screen "D_Rectangle_1" 1280x800
   TextField "Label_Static" at 6,86 size 148x16; Text 'Static'
   Rectangle "A_Range" at 158,4 size 100x50
      Appearance <- "D_Range"
   TextField "Label_A_Range" at 158,86 size 148x16; Text 'A_Range'
   Rectangle "A_Flash" at 310,4 size 100x50
      Appearance <- "D_Range"
   TextField "Label_A_Flash" at 310,86 size 148x16; Text 'A_Flash'
   Rectangle "A_Bit" at 462,4 size 100x50
      Appearance <- "D_Bool"
   TextField "Label_A_Bit" at 462,86 size 148x16; Text 'A_Bit'
   Rectangle "A_Bits" at 614,4 size 100x50
      Appearance <- "D_Bits"
   TextField "Label_A_Bits" at 614,86 size 148x16; Text 'A_Bits'
   Rectangle "V_Range" at 766,4 size 100x50
      Visibility <- "D_Range"
   TextField "Label_V_Range" at 766,86 size 148x16; Text 'V_Range'
   Rectangle "V_Bit" at 918,4 size 100x50
      Visibility <- "D_Vis"
   TextField "Label_V_Bit" at 918,86 size 148x16; Text 'V_Bit'
   Rectangle "M_H" at 1070,4 size 100x50
      HorizontalMovement <- "D_Pct"
   TextField "Label_M_H" at 1070,86 size 148x16; Text 'M_H'
   Rectangle "M_V" at 6,106 size 100x50
      VerticalMovement <- "D_Pct"
   TextField "Label_M_V" at 6,188 size 148x16; Text 'M_V'
   Rectangle "M_D" at 158,106 size 100x50
      DiagonalMovement <- "D_Pct"
   TextField "Label_M_D" at 158,188 size 148x16; Text 'M_D'
   Rectangle "M_Direct" at 310,106 size 100x50
      DirectMovement <- "D_X"
      DirectMovement <- "D_Y"
   TextField "Label_M_Direct" at 310,188 size 148x16; Text 'M_Direct'
   Rectangle "E_Range" at 462,106 size 100x50
      ObjectEnable <- "D_Range"
   TextField "Label_E_Range" at 462,188 size 148x16; Text 'E_Range'
   Rectangle "E_Bit" at 614,106 size 100x50
      ObjectEnable <- "D_En"
   TextField "Label_E_Bit" at 614,188 size 148x16; Text 'E_Bit'
   IOField "State" at 4,774 size 60x22; FormatPattern 9
      ProcessValue <- "D_State"
   Button "S1" at 70,774 size 40x22; TextOff 'S1'
      on Click: "SetS1"()
   Button "S2" at 114,774 size 40x22; TextOff 'S2'
      on Click: "SetS2"()
   Button "S3" at 158,774 size 40x22; TextOff 'S3'
      on Click: "SetS3"()
   Button "S4" at 202,774 size 40x22; TextOff 'S4'
      on Click: "SetS4"()
   Button "Next" at 1236,774 size 40x22; TextOff 'Next'
      on Click: ActivateScreen("D_TextField_1", 0)

screen "D_Slider_1" 1280x800
   Slider "Static" at 6,4 size 60x160; Caption 'SIMATIC'
   TextField "Label_Static" at 6,196 size 108x16; Text 'Static'
   Slider "A_Range" at 118,4 size 60x160; Caption 'SIMATIC'
      Appearance <- "D_Range"
   TextField "Label_A_Range" at 118,196 size 108x16; Text 'A_Range'
   Slider "A_Flash" at 230,4 size 60x160; Caption 'SIMATIC'
      Appearance <- "D_Range"
   TextField "Label_A_Flash" at 230,196 size 108x16; Text 'A_Flash'
   Slider "A_Bit" at 342,4 size 60x160; Caption 'SIMATIC'
      Appearance <- "D_Bool"
   TextField "Label_A_Bit" at 342,196 size 108x16; Text 'A_Bit'
   Slider "A_Bits" at 454,4 size 60x160; Caption 'SIMATIC'
      Appearance <- "D_Bits"
   TextField "Label_A_Bits" at 454,196 size 108x16; Text 'A_Bits'
   Slider "V_Range" at 566,4 size 60x160; Caption 'SIMATIC'
      Visibility <- "D_Range"
   TextField "Label_V_Range" at 566,196 size 108x16; Text 'V_Range'
   Slider "V_Bit" at 678,4 size 60x160; Caption 'SIMATIC'
      Visibility <- "D_Vis"
   TextField "Label_V_Bit" at 678,196 size 108x16; Text 'V_Bit'
   Slider "M_H" at 790,4 size 60x160; Caption 'SIMATIC'
      HorizontalMovement <- "D_Pct"
   TextField "Label_M_H" at 790,196 size 108x16; Text 'M_H'
   Slider "M_V" at 902,4 size 60x160; Caption 'SIMATIC'
      VerticalMovement <- "D_Pct"
   TextField "Label_M_V" at 902,196 size 108x16; Text 'M_V'
   Slider "M_D" at 1014,4 size 60x160; Caption 'SIMATIC'
      DiagonalMovement <- "D_Pct"
   TextField "Label_M_D" at 1014,196 size 108x16; Text 'M_D'
   Slider "M_Direct" at 1126,4 size 60x160; Caption 'SIMATIC'
      DirectMovement <- "D_X"
      DirectMovement <- "D_Y"
   TextField "Label_M_Direct" at 1126,196 size 108x16; Text 'M_Direct'
   Slider "E_Range" at 6,216 size 60x160; Caption 'SIMATIC'
      ObjectEnable <- "D_Range"
   TextField "Label_E_Range" at 6,408 size 108x16; Text 'E_Range'
   Slider "E_Bit" at 118,216 size 60x160; Caption 'SIMATIC'
      ObjectEnable <- "D_En"
   TextField "Label_E_Bit" at 118,408 size 108x16; Text 'E_Bit'
   Slider "PV_Pct" at 230,216 size 60x160; Caption 'SIMATIC'
      ProcessValue <- "D_Pct"
   TextField "Label_PV_Pct" at 230,408 size 108x16; Text 'PV_Pct'
   Slider "PV_Int" at 342,216 size 60x160; Caption 'SIMATIC'
      ProcessValue <- "D_Int"
   TextField "Label_PV_Int" at 342,408 size 108x16; Text 'PV_Int'
   Slider "PV_Pct_0_200" at 454,216 size 60x160; Caption 'SIMATIC'
      ProcessValue <- "D_Pct"
   TextField "Label_PV_Pct_0_200" at 454,408 size 108x16; Text 'PV_Pct_0_200'
   IOField "State" at 4,774 size 60x22; FormatPattern 9
      ProcessValue <- "D_State"
   Button "S1" at 70,774 size 40x22; TextOff 'S1'
      on Click: "SetS1"()
   Button "S2" at 114,774 size 40x22; TextOff 'S2'
      on Click: "SetS2"()
   Button "S3" at 158,774 size 40x22; TextOff 'S3'
      on Click: "SetS3"()
   Button "S4" at 202,774 size 40x22; TextOff 'S4'
      on Click: "SetS4"()
   Button "Next" at 1236,774 size 40x22; TextOff 'Next'
      on Click: ActivateScreen("D_Gauge_1", 0)

screen "D_Switch_1" 1280x800
   Switch "Static" at 6,4 size 120x40; CaptionText 'Switch'; TextOff '0'; TextOn '1'
   TextField "Label_Static" at 6,76 size 168x16; Text 'Static'
   Switch "A_Range" at 178,4 size 120x40; CaptionText 'Switch'; TextOff '0'; TextOn '1'
      Appearance <- "D_Range"
   TextField "Label_A_Range" at 178,76 size 168x16; Text 'A_Range'
   Switch "A_Flash" at 350,4 size 120x40; CaptionText 'Switch'; TextOff '0'; TextOn '1'
      Appearance <- "D_Range"
   TextField "Label_A_Flash" at 350,76 size 168x16; Text 'A_Flash'
   Switch "A_Bit" at 522,4 size 120x40; CaptionText 'Switch'; TextOff '0'; TextOn '1'
      Appearance <- "D_Bool"
   TextField "Label_A_Bit" at 522,76 size 168x16; Text 'A_Bit'
   Switch "A_Bits" at 694,4 size 120x40; CaptionText 'Switch'; TextOff '0'; TextOn '1'
      Appearance <- "D_Bits"
   TextField "Label_A_Bits" at 694,76 size 168x16; Text 'A_Bits'
   Switch "V_Range" at 866,4 size 120x40; CaptionText 'Switch'; TextOff '0'; TextOn '1'
      Visibility <- "D_Range"
   TextField "Label_V_Range" at 866,76 size 168x16; Text 'V_Range'
   Switch "V_Bit" at 1038,4 size 120x40; CaptionText 'Switch'; TextOff '0'; TextOn '1'
      Visibility <- "D_Vis"
   TextField "Label_V_Bit" at 1038,76 size 168x16; Text 'V_Bit'
   Switch "M_H" at 6,96 size 120x40; CaptionText 'Switch'; TextOff '0'; TextOn '1'
      HorizontalMovement <- "D_Pct"
   TextField "Label_M_H" at 6,168 size 168x16; Text 'M_H'
   Switch "M_V" at 178,96 size 120x40; CaptionText 'Switch'; TextOff '0'; TextOn '1'
      VerticalMovement <- "D_Pct"
   TextField "Label_M_V" at 178,168 size 168x16; Text 'M_V'
   Switch "M_D" at 350,96 size 120x40; CaptionText 'Switch'; TextOff '0'; TextOn '1'
      DiagonalMovement <- "D_Pct"
   TextField "Label_M_D" at 350,168 size 168x16; Text 'M_D'
   Switch "M_Direct" at 522,96 size 120x40; CaptionText 'Switch'; TextOff '0'; TextOn '1'
      DirectMovement <- "D_X"
      DirectMovement <- "D_Y"
   TextField "Label_M_Direct" at 522,168 size 168x16; Text 'M_Direct'
   Switch "E_Range" at 694,96 size 120x40; CaptionText 'Switch'; TextOff '0'; TextOn '1'
      ObjectEnable <- "D_Range"
   TextField "Label_E_Range" at 694,168 size 168x16; Text 'E_Range'
   Switch "E_Bit" at 866,96 size 120x40; CaptionText 'Switch'; TextOff '0'; TextOn '1'
      ObjectEnable <- "D_En"
   TextField "Label_E_Bit" at 866,168 size 168x16; Text 'E_Bit'
   Switch "PV_Bool" at 1038,96 size 120x40; CaptionText 'Switch'; TextOff '0'; TextOn '1'
      ProcessValue <- "D_Bool"
   TextField "Label_PV_Bool" at 1038,168 size 168x16; Text 'PV_Bool'
   IOField "State" at 4,774 size 60x22; FormatPattern 9
      ProcessValue <- "D_State"
   Button "S1" at 70,774 size 40x22; TextOff 'S1'
      on Click: "SetS1"()
   Button "S2" at 114,774 size 40x22; TextOff 'S2'
      on Click: "SetS2"()
   Button "S3" at 158,774 size 40x22; TextOff 'S3'
      on Click: "SetS3"()
   Button "S4" at 202,774 size 40x22; TextOff 'S4'
      on Click: "SetS4"()
   Button "Next" at 1236,774 size 40x22; TextOff 'Next'
      on Click: ActivateScreen("D_SymbolLibrary_1", 0)

screen "D_SymbolicIOField_1" 1280x800
   SymbolicIOField "Static" at 6,4 size 120x30; TextOff '0'; TextOn '1'
   TextField "Label_Static" at 6,66 size 168x16; Text 'Static'
   SymbolicIOField "A_Range" at 178,4 size 120x30; TextOff '0'; TextOn '1'
      Appearance <- "D_Range"
   TextField "Label_A_Range" at 178,66 size 168x16; Text 'A_Range'
   SymbolicIOField "A_Flash" at 350,4 size 120x30; TextOff '0'; TextOn '1'
      Appearance <- "D_Range"
   TextField "Label_A_Flash" at 350,66 size 168x16; Text 'A_Flash'
   SymbolicIOField "A_Bit" at 522,4 size 120x30; TextOff '0'; TextOn '1'
      Appearance <- "D_Bool"
   TextField "Label_A_Bit" at 522,66 size 168x16; Text 'A_Bit'
   SymbolicIOField "A_Bits" at 694,4 size 120x30; TextOff '0'; TextOn '1'
      Appearance <- "D_Bits"
   TextField "Label_A_Bits" at 694,66 size 168x16; Text 'A_Bits'
   SymbolicIOField "V_Range" at 866,4 size 120x30; TextOff '0'; TextOn '1'
      Visibility <- "D_Range"
   TextField "Label_V_Range" at 866,66 size 168x16; Text 'V_Range'
   SymbolicIOField "V_Bit" at 1038,4 size 120x30; TextOff '0'; TextOn '1'
      Visibility <- "D_Vis"
   TextField "Label_V_Bit" at 1038,66 size 168x16; Text 'V_Bit'
   SymbolicIOField "M_H" at 6,86 size 120x30; TextOff '0'; TextOn '1'
      HorizontalMovement <- "D_Pct"
   TextField "Label_M_H" at 6,148 size 168x16; Text 'M_H'
   SymbolicIOField "M_V" at 178,86 size 120x30; TextOff '0'; TextOn '1'
      VerticalMovement <- "D_Pct"
   TextField "Label_M_V" at 178,148 size 168x16; Text 'M_V'
   SymbolicIOField "M_D" at 350,86 size 120x30; TextOff '0'; TextOn '1'
      DiagonalMovement <- "D_Pct"
   TextField "Label_M_D" at 350,148 size 168x16; Text 'M_D'
   SymbolicIOField "M_Direct" at 522,86 size 120x30; TextOff '0'; TextOn '1'
      DirectMovement <- "D_X"
      DirectMovement <- "D_Y"
   TextField "Label_M_Direct" at 522,148 size 168x16; Text 'M_Direct'
   SymbolicIOField "E_Range" at 694,86 size 120x30; TextOff '0'; TextOn '1'
      ObjectEnable <- "D_Range"
   TextField "Label_E_Range" at 694,148 size 168x16; Text 'E_Range'
   SymbolicIOField "E_Bit" at 866,86 size 120x30; TextOff '0'; TextOn '1'
      ObjectEnable <- "D_En"
   TextField "Label_E_Bit" at 866,148 size 168x16; Text 'E_Bit'
   SymbolicIOField "PV_TL_Value" at 1038,86 size 120x30; TextOff '0'; TextOn '1'; TextList "TL_Value"
      ProcessValue <- "D_TL"
   TextField "Label_PV_TL_Value" at 1038,148 size 168x16; Text 'PV_TL_Value'
   SymbolicIOField "PV_TL_Bit" at 6,168 size 120x30; TextOff '0'; TextOn '1'; TextList "TL_Bit"
      ProcessValue <- "D_Bool"
   TextField "Label_PV_TL_Bit" at 6,230 size 168x16; Text 'PV_TL_Bit'
   SymbolicIOField "PV_TL_BitNo" at 178,168 size 120x30; TextOff '0'; TextOn '1'; TextList "TL_BitNo"
      ProcessValue <- "D_Bits"
   TextField "Label_PV_TL_BitNo" at 178,230 size 168x16; Text 'PV_TL_BitNo'
   IOField "State" at 4,774 size 60x22; FormatPattern 9
      ProcessValue <- "D_State"
   Button "S1" at 70,774 size 40x22; TextOff 'S1'
      on Click: "SetS1"()
   Button "S2" at 114,774 size 40x22; TextOff 'S2'
      on Click: "SetS2"()
   Button "S3" at 158,774 size 40x22; TextOff 'S3'
      on Click: "SetS3"()
   Button "S4" at 202,774 size 40x22; TextOff 'S4'
      on Click: "SetS4"()
   Button "Next" at 1236,774 size 40x22; TextOff 'Next'
      on Click: ActivateScreen("D_GraphicIOField_1", 0)

screen "D_SymbolLibrary_1" 1280x800
   SymbolLibrary "Static" at 6,4 size 60x60
   TextField "Label_Static" at 6,96 size 108x16; Text 'Static'
   SymbolLibrary "A_Range" at 118,4 size 60x60
      Appearance <- "D_Range"
   TextField "Label_A_Range" at 118,96 size 108x16; Text 'A_Range'
   SymbolLibrary "A_Flash" at 230,4 size 60x60
      Appearance <- "D_Range"
   TextField "Label_A_Flash" at 230,96 size 108x16; Text 'A_Flash'
   SymbolLibrary "A_Bit" at 342,4 size 60x60
      Appearance <- "D_Bool"
   TextField "Label_A_Bit" at 342,96 size 108x16; Text 'A_Bit'
   SymbolLibrary "A_Bits" at 454,4 size 60x60
      Appearance <- "D_Bits"
   TextField "Label_A_Bits" at 454,96 size 108x16; Text 'A_Bits'
   SymbolLibrary "V_Range" at 566,4 size 60x60
      Visibility <- "D_Range"
   TextField "Label_V_Range" at 566,96 size 108x16; Text 'V_Range'
   SymbolLibrary "V_Bit" at 678,4 size 60x60
      Visibility <- "D_Vis"
   TextField "Label_V_Bit" at 678,96 size 108x16; Text 'V_Bit'
   SymbolLibrary "M_H" at 790,4 size 60x60
      HorizontalMovement <- "D_Pct"
   TextField "Label_M_H" at 790,96 size 108x16; Text 'M_H'
   SymbolLibrary "M_V" at 902,4 size 60x60
      VerticalMovement <- "D_Pct"
   TextField "Label_M_V" at 902,96 size 108x16; Text 'M_V'
   SymbolLibrary "M_D" at 1014,4 size 60x60
      DiagonalMovement <- "D_Pct"
   TextField "Label_M_D" at 1014,96 size 108x16; Text 'M_D'
   SymbolLibrary "M_Direct" at 1126,4 size 60x60
      DirectMovement <- "D_X"
      DirectMovement <- "D_Y"
   TextField "Label_M_Direct" at 1126,96 size 108x16; Text 'M_Direct'
   SymbolLibrary "E_Range" at 6,116 size 60x60
      ObjectEnable <- "D_Range"
   TextField "Label_E_Range" at 6,208 size 108x16; Text 'E_Range'
   SymbolLibrary "E_Bit" at 118,116 size 60x60
      ObjectEnable <- "D_En"
   TextField "Label_E_Bit" at 118,208 size 108x16; Text 'E_Bit'
   SymbolLibrary "PV_Pct" at 230,116 size 60x60
      ProcessValue <- "D_Pct"
   TextField "Label_PV_Pct" at 230,208 size 108x16; Text 'PV_Pct'
   IOField "State" at 4,774 size 60x22; FormatPattern 9
      ProcessValue <- "D_State"
   Button "S1" at 70,774 size 40x22; TextOff 'S1'
      on Click: "SetS1"()
   Button "S2" at 114,774 size 40x22; TextOff 'S2'
      on Click: "SetS2"()
   Button "S3" at 158,774 size 40x22; TextOff 'S3'
      on Click: "SetS3"()
   Button "S4" at 202,774 size 40x22; TextOff 'S4'
      on Click: "SetS4"()
   Button "Next" at 1236,774 size 40x22; TextOff 'Next'
      on Click: ActivateScreen("D_Slider_1", 0)

screen "D_TextField_1" 1280x800
   TextField "Static" at 6,4 size 100x30; Text 'Text'
   TextField "Label_Static" at 6,66 size 148x16; Text 'Static'
   TextField "A_Range" at 158,4 size 100x30; Text 'Text'
      Appearance <- "D_Range"
   TextField "Label_A_Range" at 158,66 size 148x16; Text 'A_Range'
   TextField "A_Flash" at 310,4 size 100x30; Text 'Text'
      Appearance <- "D_Range"
   TextField "Label_A_Flash" at 310,66 size 148x16; Text 'A_Flash'
   TextField "A_Bit" at 462,4 size 100x30; Text 'Text'
      Appearance <- "D_Bool"
   TextField "Label_A_Bit" at 462,66 size 148x16; Text 'A_Bit'
   TextField "A_Bits" at 614,4 size 100x30; Text 'Text'
      Appearance <- "D_Bits"
   TextField "Label_A_Bits" at 614,66 size 148x16; Text 'A_Bits'
   TextField "V_Range" at 766,4 size 100x30; Text 'Text'
      Visibility <- "D_Range"
   TextField "Label_V_Range" at 766,66 size 148x16; Text 'V_Range'
   TextField "V_Bit" at 918,4 size 100x30; Text 'Text'
      Visibility <- "D_Vis"
   TextField "Label_V_Bit" at 918,66 size 148x16; Text 'V_Bit'
   TextField "M_H" at 1070,4 size 100x30; Text 'Text'
      HorizontalMovement <- "D_Pct"
   TextField "Label_M_H" at 1070,66 size 148x16; Text 'M_H'
   TextField "M_V" at 6,86 size 100x30; Text 'Text'
      VerticalMovement <- "D_Pct"
   TextField "Label_M_V" at 6,148 size 148x16; Text 'M_V'
   TextField "M_D" at 158,86 size 100x30; Text 'Text'
      DiagonalMovement <- "D_Pct"
   TextField "Label_M_D" at 158,148 size 148x16; Text 'M_D'
   TextField "M_Direct" at 310,86 size 100x30; Text 'Text'
      DirectMovement <- "D_X"
      DirectMovement <- "D_Y"
   TextField "Label_M_Direct" at 310,148 size 148x16; Text 'M_Direct'
   TextField "E_Range" at 462,86 size 100x30; Text 'Text'
      ObjectEnable <- "D_Range"
   TextField "Label_E_Range" at 462,148 size 148x16; Text 'E_Range'
   TextField "E_Bit" at 614,86 size 100x30; Text 'Text'
      ObjectEnable <- "D_En"
   TextField "Label_E_Bit" at 614,148 size 148x16; Text 'E_Bit'
   IOField "State" at 4,774 size 60x22; FormatPattern 9
      ProcessValue <- "D_State"
   Button "S1" at 70,774 size 40x22; TextOff 'S1'
      on Click: "SetS1"()
   Button "S2" at 114,774 size 40x22; TextOff 'S2'
      on Click: "SetS2"()
   Button "S3" at 158,774 size 40x22; TextOff 'S3'
      on Click: "SetS3"()
   Button "S4" at 202,774 size 40x22; TextOff 'S4'
      on Click: "SetS4"()
   Button "Next" at 1236,774 size 40x22; TextOff 'Next'
      on Click: ActivateScreen("D_GraphicView_1", 0)

VB script "SetS1"
   SmartTags("D_State") = 1
   SmartTags("D_Bool") = False
   SmartTags("D_SInt") = -128
   SmartTags("D_Int") = -32768
   SmartTags("D_DInt") = -2147483648
   SmartTags("D_USInt") = 0
   SmartTags("D_UInt") = 0
   SmartTags("D_UDInt") = 0
   SmartTags("D_Real") = -999.999
   SmartTags("D_LReal") = -0.00000015
   SmartTags("D_String") = ""
   SmartTags("D_DateTime") = DateSerial(1990, 1, 1) + TimeSerial(0, 0, 0)
   SmartTags("D_Pct") = 0
   SmartTags("D_Range") = 5
   SmartTags("D_Bits") = 1
   SmartTags("D_Vis") = False
   SmartTags("D_En") = False
   SmartTags("D_X") = 10
   SmartTags("D_Y") = 10
   SmartTags("D_Max") = 100
   SmartTags("D_Min") = 0
   SmartTags("D_TL") = -5
   SmartTags("D_BarR") = -5

VB script "SetS2"
   SmartTags("D_State") = 2
   SmartTags("D_Bool") = True
   SmartTags("D_SInt") = 12
   SmartTags("D_Int") = 1234
   SmartTags("D_DInt") = 123456
   SmartTags("D_USInt") = 200
   SmartTags("D_UInt") = 40000
   SmartTags("D_UDInt") = 3000000000
   SmartTags("D_Real") = 3.14159
   SmartTags("D_LReal") = 2.718281828
   SmartTags("D_String") = "Hello World"
   SmartTags("D_DateTime") = DateSerial(2026, 11, 22) + TimeSerial(13, 45, 30)
   SmartTags("D_Pct") = 50
   SmartTags("D_Range") = 25
   SmartTags("D_Bits") = 2
   SmartTags("D_Vis") = True
   SmartTags("D_En") = True
   SmartTags("D_X") = 320
   SmartTags("D_Y") = 200
   SmartTags("D_Max") = 200
   SmartTags("D_Min") = -100
   SmartTags("D_TL") = 5
   SmartTags("D_BarR") = 0

VB script "SetS3"
   SmartTags("D_State") = 3
   SmartTags("D_Bool") = True
   SmartTags("D_SInt") = 127
   SmartTags("D_Int") = 32767
   SmartTags("D_DInt") = 2147483647
   SmartTags("D_USInt") = 255
   SmartTags("D_UInt") = 65535
   SmartTags("D_UDInt") = 4294967295
   SmartTags("D_Real") = 123456.789
   SmartTags("D_LReal") = 1E+300
   SmartTags("D_String") = "Ünïcödé äöüß ÄÖÜ € – long text that is wider than the field 0123456789 ABCDEFGHIJ"
   SmartTags("D_DateTime") = DateSerial(2099, 12, 31) + TimeSerial(23, 59, 59)
   SmartTags("D_Pct") = 100
   SmartTags("D_Range") = 75
   SmartTags("D_Bits") = 4
   SmartTags("D_Vis") = True
   SmartTags("D_En") = False
   SmartTags("D_X") = 853
   SmartTags("D_Y") = 400
   SmartTags("D_Max") = 50
   SmartTags("D_Min") = -50
   SmartTags("D_TL") = 10
   SmartTags("D_BarR") = 5

VB script "SetS4"
   SmartTags("D_State") = 4
   SmartTags("D_Bool") = False
   SmartTags("D_SInt") = -1
   SmartTags("D_Int") = -1
   SmartTags("D_DInt") = 0
   SmartTags("D_USInt") = 1
   SmartTags("D_UInt") = 1
   SmartTags("D_UDInt") = 1
   SmartTags("D_Real") = 0.0005
   SmartTags("D_LReal") = -0.0
   SmartTags("D_String") = "äöü ÄÖÜ ß"
   SmartTags("D_DateTime") = DateSerial(1970, 1, 1) + TimeSerial(0, 0, 0)
   SmartTags("D_Pct") = 150
   SmartTags("D_Range") = 200
   SmartTags("D_Bits") = 9
   SmartTags("D_Vis") = False
   SmartTags("D_En") = True
   SmartTags("D_X") = -20
   SmartTags("D_Y") = 0
   SmartTags("D_Max") = 100
   SmartTags("D_Min") = 0
   SmartTags("D_TL") = 50
   SmartTags("D_BarR") = 2.5
*)